{attribute 'qualified_only'}
VAR_GLOBAL
	command : SimulatorCommand;
	feedback : SimulatorFeedback;
	scan : LaserScan;
END_VAR

(* stored: Version 1.1.0.1, ProductVersion 3.1.4026.12
   GVL SimulatorIo: Id {9fa4ee25-d7a0-5946-92a6-d883b06d34b4} *)
